# EPICS substitutions: iocs/motor/smartmotor-ioc/db/SmartMotor.substitutions
# C's iocSmartMotor SmartMotor.substitutions, P and C from st.cmd. Signal S
# is chain axis S; VELO and ACCL feed V= and A=.
file "$(MOTOR)/db/motor.db"
{
pattern
{N,  M,        DTYP,          S,  DESC,          EGU,      DIR,  VELO,  VBAS,  ACCL,  BDST,  BVEL,  BACC,  MRES,  PREC,  DHLM,  DLLM,  INIT}
{1,  "m$(N)",  "SmartMotor",  0,  "motor $(N)",  degrees,  Pos,  1,     .1,    .2,    0,     1,     .2,    0.01,  5,     100,   -100,  ""}
}
